Fanuc KAREL source: ko00064.KL

PROGRAM KO00064
%STACKSIZE=65535
%PRIORITY=65535
%NOLOCKGROUP
VAR
P1 : XYZWPR
P2 : JOINTPOS9
F : BOOLEAN
OUT : JOINTPOS9
BEGIN
F=TRUE
-- UNSAFE_SOURCE_IR line 11: CALL_RESULT MIRROR(convert_xyzwpr_to_xyzwprext(P1), convert_jointpos9_to_position(P2), F)
END KO00064
